(* CODESYS project PLC_PRG.xml

Project tree, tasks and I/O mapping:
  program PLC_PRG [CFC]
*)

// PLC_PRG
// The program activates or deactivates the cooling compressor depending on the 
// deviaton of the actual temperature from the septpoint temperature (with a hysteresis)

// TRUE or FALSE of the cooling compresseor is transfered to the signal processing.
PROGRAM PLC_PRG
VAR
	SR_0: SR;
	Hysteresis: REAL:=1.0;
END_VAR

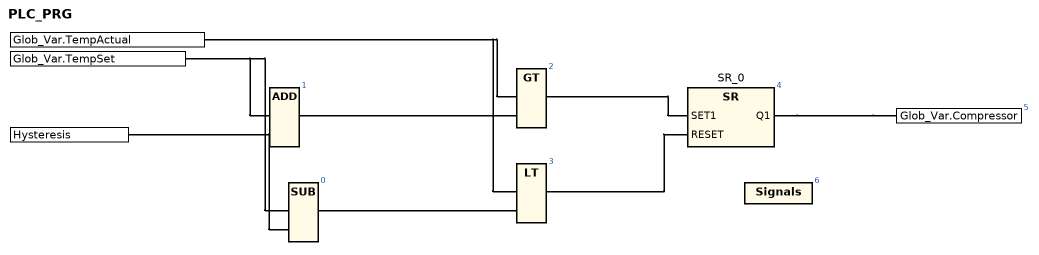
// note: 1 stored wires end on pins the file does not list and are not shown
SR_0(SET1 := Glob_Var.TempActual > Glob_Var.TempSet + Hysteresis, RESET := Glob_Var.TempActual < Glob_Var.TempSet - Hysteresis); // SR
Glob_Var.Compressor := SR_0.Q1;
Signals();

END_PROGRAM
